FUNCTION F_RealToBitDword : DWORD
VAR_INPUT
	rIn : REAL;
END_VAR
VAR
	pt : POINTER TO DWORD;
END_VAR

pt := ADR(rIn);
F_RealToBitDword := pt^;

END_FUNCTION

(* stored: Version 1.1.0.1, ProductVersion 3.1.4024.15
   POU F_RealToBitDword: Id {e777d8b4-422e-4dcb-8434-6fc347c18a79}, SpecialFunc None *)
